// TIA Portal V21 export
// export: Created 2026-10-23T20:44:33.4914774Z, ExportSetting WithDefaults, DisplayName Totally Integrated Automation Portal, DisplayVersion V21 Update 1, DisplayName SINAMICS Startdrive Advanced, DisplayVersion V21 HF2, DisplayName SINAMICS Startdrive G110M, G120, G120C, G120D, G120P, G115D, DisplayVersion V21 HF2, DisplayName SINAMICS Startdrive G130, G150, S120, S150, G200, G220, S200, S210, S220, Innomotics MVD, DisplayVersion V21 HF2, DisplayName STEP 7 Professional, DisplayVersion V21 Update 1, DisplayName STEP 7 Safety, DisplayVersion V21, DisplayName Tech WebApplication, DisplayVersion V21, DisplayName WinCC Basic/Comfort/Advanced, DisplayVersion V21 Update 1, DisplayName WinCC Unified, DisplayVersion V21 Update 1
FUNCTION "FC_FillHelper" : Real   // FC7, SCL
TITLE = Volume from raw flow
VERSION : 0.1
// Unpublished helper of the filling unit
// stored: Access Unpublished, AutoNumber true, IsIECCheckEnabled false, Namespace Filling, SetENOAutomatically false, UDAEnableTagReadback false
   VAR_INPUT
      RawFlow : Int;   // Raw flow value
      Factor : Real;   // Litres per raw unit
   END_VAR
BEGIN

       #FC_FillHelper := INT_TO_REAL(#RawFlow) * #Factor;
END_FUNCTION
